Fanuc KAREL source: KA00063.KL

PROGRAM KA00063
%NOLOCKGROUP
VAR
  SRC: XYZWPR
  DST: BOOLEAN
BEGIN
  SRC.X = 1.0
  DST = SRC
END KA00063
